{region 'Documentation'}
(*!
<summary>Supplies controlled parent identity for Assertion initialization tests.</summary>
<description>
Only Name is consumed by the subject. SetIdentity deliberately admits malformed names
to exercise the subject boundary. This local mock is never scheduled as a Test Case.
</description>
*)
{endregion}
FUNCTION_BLOCK AssertionParentIdentity EXTENDS TestCaseMock

SUPER^();

{region 'Documentation'}
(*!
<summary>Sets the parent name before the subject reads it; no lifecycle work.</summary>
*)
{endregion}
METHOD PUBLIC SetIdentity
VAR_INPUT
    Value : STRING(GVL_Constants.NameLength); //! Identity-only parent name retained for isolated Assertion initialization.
END_VAR
FName := Value;
END_METHOD

END_FUNCTION_BLOCK

(* stored: Version 1.1.0.1
   POU AssertionParentIdentity: Id {d80bd656-9f6b-4065-bc47-a98ab5309d3f}, SpecialFunc None
   Folder Internal: Id {7c4afd2f-6b20-4a4b-8263-a776d9905dba}
   Method SetIdentity: Id {c6037e91-be61-43eb-a0ad-67cb71204722} *)
